(* IEC 61131-3 sources: codesys-framework/txt/application/WeVe Core (library)/00 Application, 1 file *)

(* ---- FB_Application.pou.st ---- *)
FUNCTION_BLOCK ABSTRACT FB_Application IMPLEMENTS I_Application
VAR_INPUT
END_VAR
VAR_OUTPUT
END_VAR
VAR
END_VAR

// --- BEGIN IMPLEMENTATION ---
